(* IEC 61131-3 sources: Versio-VersionControlSystem/fixtures/projects/TC3_PlcSample_reStrText/TC3_PlcSample_reStrText/LibraryDocumentationSample Project/LibPOUs/B_DocuElements/Tables, 4 files *)

(* ---- FB_Libdoc_CSVTable.st ---- *)
(*
.. csv-table:: Property list
   :header: "Items", "Property 1", "Property 2", "Property 3"
   :widths: 10, 15, 15, 15

   "Item 1", 1.67, angular, red
   "Item 2", "not specified", round, blue

|

.. csv-table:: Property list
   :header-rows: 1
   :widths: 10, 15, 15, 15

   "Items", "Property 1", "Property 2", "Property 3"
   "Item 1", 1.67, angular, red
   "Item 2", "not specified", round, blue
*)

FUNCTION_BLOCK FB_Libdoc_CSVTable
VAR_INPUT
    nVarA : INT;
    nVarB : INT;
END_VAR
VAR_OUTPUT
    nSum : INT;
END_VAR
VAR
END_VAR

(* ---- FB_Libdoc_GridTable.st ---- *)
(*
+------------------------+------------+----------+----------+
| Header row, column 1   | Header 2   | Header 3 | Header 4 |
| (header rows optional) |            |          |          |
+========================+============+==========+==========+
| body row 1, column 1   | column 2   | column 3 | column 4 |
+------------------------+------------+----------+----------+
| body row 2             | Cells may span columns.          |
+------------------------+------------+---------------------+
| body row 3             | Cells may  | - Table cells       |
+------------------------+ span rows. | - contain           |
| body row 4             |            | - body elements.    |
+------------------------+------------+---------------------+
*)

FUNCTION_BLOCK FB_Libdoc_GridTable
VAR_INPUT
    nVarA : INT;
    nVarB : INT;
END_VAR
VAR_OUTPUT
    nSum : INT;
END_VAR
VAR
END_VAR

(* ---- FB_Libdoc_ListTable.st ---- *)
(*
.. list-table:: Property list
    :widths: 50 50 50
    :header-rows: 1

    * - Items
      - Property 1
      - Property 2
    * - Item 1
      - angular
      - red
    * - Item 2
      - round
      - blue
*)

FUNCTION_BLOCK FB_Libdoc_ListTable
VAR_INPUT
    nVarA : INT;
    nVarB : INT;
END_VAR
VAR_OUTPUT
    nSum : INT;
END_VAR
VAR
END_VAR

(* ---- FB_Libdoc_SimpleTables.st ---- *)
(*
=====  =====  =======
  A      B    A and B
=====  =====  =======
False  False  False
True   False  False
False  True   False
True   True   True
=====  =====  =======

|

=====  =====  ======
   Inputs     Output
------------  ------
  A      B    A or B
=====  =====  ======
False  False  False
True   False  True
False  True   True
True   True   True
=====  =====  ======

|

=====  =====  ======
   Inputs     Output
------------  ------
  A      B    A or B
=====  =====  ======
False  False  False
       False  True
False  True   True
True   True   True
=====  =====  ======

|

=====  =====
Col 1  Col 2
=====  =====
1      Second column of row 1.
2      Second column of row 2.
       Second line of paragraph.
3      Second column of row 2.

       Second line of paragraph
4      - Second column of row 3.

       - Second item in bullet
         list (row 4, column 2).
\      Row 5; column 1 will be empty.
=====  =====
*)

FUNCTION_BLOCK FB_Libdoc_SimpleTables
VAR_INPUT
    nVarA : INT;
    nVarB : INT;
END_VAR
VAR_OUTPUT
    nSum : INT;
END_VAR
VAR
END_VAR
